(* IEC 61131-3 sources: Lasal-MCP/examples/SampleSource/LASALScreenAdvancedSolution/LASALScreenAdvancedSolution/LASALScreenAdvacnedSolution/Stations/MachineControl/MachineControl/Class/VaranManager (part 5) *)

    DPRAM_Used.Total              += sizeof(LSL_VARANFRAMEPAYLOADMOVEHEADER) + 1 + sizeof(LSL_VARANFRAMEMOVEWRITEPAYLOAD);  // Header + Read Statusbyte + Write Payload
    DPRAM_Used_Payload.Total      += 1 + sizeof(LSL_VARANFRAMEMOVEWRITEPAYLOAD);  // Read Statusbyte + Write Payload
    DOCounter.Total               += 1;
  end_if;

END_FUNCTION

FUNCTION VaranManager::GetDataPointers
  VAR_INPUT
    ud_hDoHandle 	: UDINT;
    pp_ReadData 	: ^pVoid;
    pp_WriteData 	: ^pVoid;
  END_VAR
  VAR_OUTPUT
    sd_retval 	  : DINT;
  END_VAR

#ifdef VM_DEBUG_PAYLOAD
  if b_PayloadSupport = false then
    // This method is not suppored without payload
    ((0)$^USINT)^ := 0;
  end_if;
#endif

  // if there is no VARAN Interface available, we would crash at the call
  if pMultiVaran = NIL then
    sd_retval := VARANMANAGER_DRIVER_NOT_EXISTS;
    return;
  end_if;

  sd_retval :=  MULTI_VARAN_iGetDataPointers( hDoHandle   := ud_hDoHandle
                                            , ppvReadData := pp_ReadData
                                            , ppvWriteData:= pp_WriteData
                                            );

END_FUNCTION

FUNCTION VaranManager::GetModuleHandle
  VAR_INPUT
    p_us_PositionInfo 	: ^USINT;
    p_ud_ModuleHandle 	: ^UDINT;
  END_VAR
  VAR_OUTPUT
    sd_retval 	        : DINT;
  END_VAR

  // if there is no VARAN Interface available, we would crash at the call
  if pMultiVaran = NIL then
    sd_retval := VARANMANAGER_DRIVER_NOT_EXISTS;
    return;
  end_if;

  sd_retval := MULTI_VARAN_iGetNodeHandle(  udManagerNumber := VaranManagerNr
                                          , pszHardwarePath := p_us_PositionInfo
                                          , phNodeHandle    := p_ud_ModuleHandle
                                          );

END_FUNCTION

FUNCTION VaranManager::AddObjectCallback
	VAR_INPUT
		p_us_position_info 	: ^USINT;
		ud_action_ptr 	    : UDINT;
		ud_thisp 	          : UDINT;
		sd_required 	      : DINT;
	END_VAR
	VAR_OUTPUT
		sd_retval 	        : DINT;
	END_VAR
  VAR
    ud_NodeHandle       : UDINT;
  END_VAR

  if State = _NoVaranInterface then
    sd_retval := -100;
    return;
  end_if;
  //get right required flag
  if ( sd_required ) then
    sd_required := VARAN_DEVICE_REQUIRED;
  else
    sd_required := VARAN_DEVICE_DEFAULT;
  end_if;

  if b_PayloadSupport &
       pMultiVaran^.udVersion >= VM_MULTIVARAN_VERSION_FULL_PAYLOAD_AVAILABLE  then
    sd_retval := MULTI_VARAN_iGetNodeHandle ( udManagerNumber := VaranManagerNr
                                            , pszHardwarePath := p_us_position_info
                                            , phNodeHandle    := #ud_NodeHandle
                                            );

    if sd_retval <> VARANMANAGER_OK then
      return;
    end_if;

    //call OS - function to set callback
    sd_retval := MULTI_VARAN_iSetApplicationCallback( hNodeHandle           := ud_NodeHandle
                                                    , pfApplicationCallback := ud_action_ptr$pvoid
                                                    , pvUserData            := ud_thisp$pvoid
                                                    , udRequired            := sd_required$UDINT
                                                    );

  elsif pVaran then

    //call OS - function to set callback
    sd_retval := VARAN_iSetObjectCallback	( uiManager   := VaranManagerNr
                                          , pucNode     := p_us_position_info
                                          , uiCallback  := ud_action_ptr
                                          , uiThis      := ud_thisp
                                          , uiRequired  := sd_required$UDINT
                                          );
  end_if;

  //look for an error
  if ( sd_retval <> VARANMANAGER_OK ) then
    s_ErrorVaranManager.f_SetObjectCallback := SetVaranDOError	( sd_Error 		  := sd_retval
                                                                , b_manager_off	:= TRUE
                                                                , b_log			    := TRUE
                                                                );
  end_if;

END_FUNCTION

FUNCTION VaranManager::GetSPIDataFromID
	VAR_INPUT
		p_us_position_info 	: ^USINT;
		udListID 	          : UDINT;
		pData 	            : ^CHAR;
		udRequDataLength 	  : UDINT;
		pIDHeader 	        : ^t_s_SPIListHeader;
		udOffset 	          : UDINT;(* := 16#00 *)
	END_VAR
	VAR_OUTPUT
		sd_retval 	        : DINT;
	END_VAR
  VAR
    BaseListAddress     : UDINT;
    a_data              : ARRAY[0..31] OF UDINT;
  END_VAR

  if p_us_position_info & pData & udRequDataLength > 0 then

    //check OS version
    if ( _RTOSVersion < VM_SPI_OS_VERSION ) then
      // access of SPI flash not possible
      sd_retval := -2;
      return;
    end_if;

    // check if list is available and get size and offset in SPI flash
    if ( SearchSPIList(p_us_position_info, udListID, #BaseListAddress) <> VARANMANAGER_OK ) then
      sd_retval := -3;
      return;
    end_if;

    //read header of list
    sd_retval := ReadSPIDataComfort(p_us_position_info  := p_us_position_info,
                                    ud_offset           := BaseListAddress,
                                    ud_length	          := sizeof(t_s_SPIListHeader),
                                    p_data	            := ( #a_data )$^USINT
                                    );

    _memcpy(ptr1:=pIDHeader, ptr2:=#a_data[0], cntr:=sizeof(t_s_SPIListHeader));

    //look for an error and check if length is > 0
    if ( sd_retval <> VARANMANAGER_OK ) | ( a_data[ 2 ] = 0 ) then
      sd_retval := -4;
      return;
    end_if;

    //read the whole serial number string
    sd_retval := ReadSPIDataComfort( p_us_position_info := p_us_position_info,
                                     ud_offset	        := BaseListAddress + sizeof(t_s_SPIListHeader) + udOffset,  //+12 ist List Header
                                     ud_length	        := udRequDataLength,
                                     p_data		          := pData
                                    );

    //look for an error
    if ( sd_retval <> VARANMANAGER_OK ) then
      sd_retval := -5;
      return;
    end_if;
  else
    // invalid parameters
    sd_retval := -1;
  end_if;

END_FUNCTION

FUNCTION GLOBAL VaranManager::RaiseManagerError
	VAR_INPUT
		udReason 	: UDINT;
	END_VAR

  State := udReason$t_e_VaranErrors;

  if b_PayloadSupport & pMultiVaran^.udVersion >= VM_MULTIVARAN_VERSION_FULL_PAYLOAD_AVAILABLE  then
    MULTI_VARAN_iReportVaranError( diErrorNumber := udReason$DINT
                                 , hErrorNode    := vmNodeHandle
                                 );

  elsif pVaran & (pVaran^.udVersion >= 16#00001104 ) then
    VARAN_iSetManagerError( VaranManagerNr, udReason );
  end_if;

END_FUNCTION
